// TIA Portal V21 export
// export: Created 2026-10-09T20:27:00.7380612Z, ExportSetting WithDefaults, DisplayName Totally Integrated Automation Portal, DisplayVersion V21, DisplayName STEP 7 Professional, DisplayVersion V21, DisplayName STEP 7 Safety, DisplayVersion V21, DisplayName Tech WebApplication, DisplayVersion V21, DisplayName WinCC Basic/Comfort/Advanced, DisplayVersion V21, DisplayName WinCC Unified, DisplayVersion V21
FUNCTION_BLOCK "FB_2_Filling"   // FB3, FBD
TITLE = Filling process
{ S7_Optimized_Access := 'TRUE' }
VERSION : 0.1
// stored: AutoNumber true, IsIECCheckEnabled false, IsRetainMemResEnabled false, MemoryReserve 100, SetENOAutomatically false, UDAEnableTagReadback false
   VAR_INPUT
      externalSignals : "typeSignals";   // signals from external model
   END_VAR
   VAR_IN_OUT
      model : "typeModel";   // model parameter
      operate : "typeOperate";   // application operation
      signals : "typeSignals";   // current signals from tank
      process : "typeProcess";   // current process information
      appSignals : "typeApp";
      hmiSignals : "typeHmi";
      errors : "typeError";   // error information
   END_VAR
   VAR
      statShiftingBottle : Bool;
      statShiftingTrigger : Bool;
      statShiftingTimer : Int;
      statHmiBottleLevel : Real;   // parameter for HMI to show current bottle level
      statHmiDoShift : Bool;   // trigger for HMI to shift bottles
      statHmiFaultyBottle : Bool;   // trigger for HMI for faulty bottle
      statBatchIdOld { ExternalAccessible := 'False'; ExternalVisible := 'False'; ExternalWritable := 'False'} : UDInt := 0;   // helper when batchID changed
      statFillingTankTrigger : Bool;
      statStartCounter { ExternalAccessible := 'False'; ExternalVisible := 'False'; ExternalWritable := 'False'} : Bool;
      statProducedStart { ExternalAccessible := 'False'; ExternalVisible := 'False'; ExternalWritable := 'False'} : UDInt;
      statProducedEnd { ExternalAccessible := 'False'; ExternalVisible := 'False'; ExternalWritable := 'False'} : UDInt;
      statSizeBatchID : USInt;
      statSizeNumberProduced : USInt;
      statStringBatchID : String;
      statStringProductID : String;
   END_VAR
   VAR_TEMP
      tempBottleMaxLevel : Real;
      tempTimerFinished : Bool;
      tempTimeOutput : Time;
      tempCurrentTime : DTL;
      tempTimeRet : Int;
   END_VAR
   VAR_TEMP   // added for the SCL form of the ladder/FBD networks
      _w1 : Bool;
      _w2 : Bool;
   END_VAR
BEGIN

REGION Network 1: Calculation of params
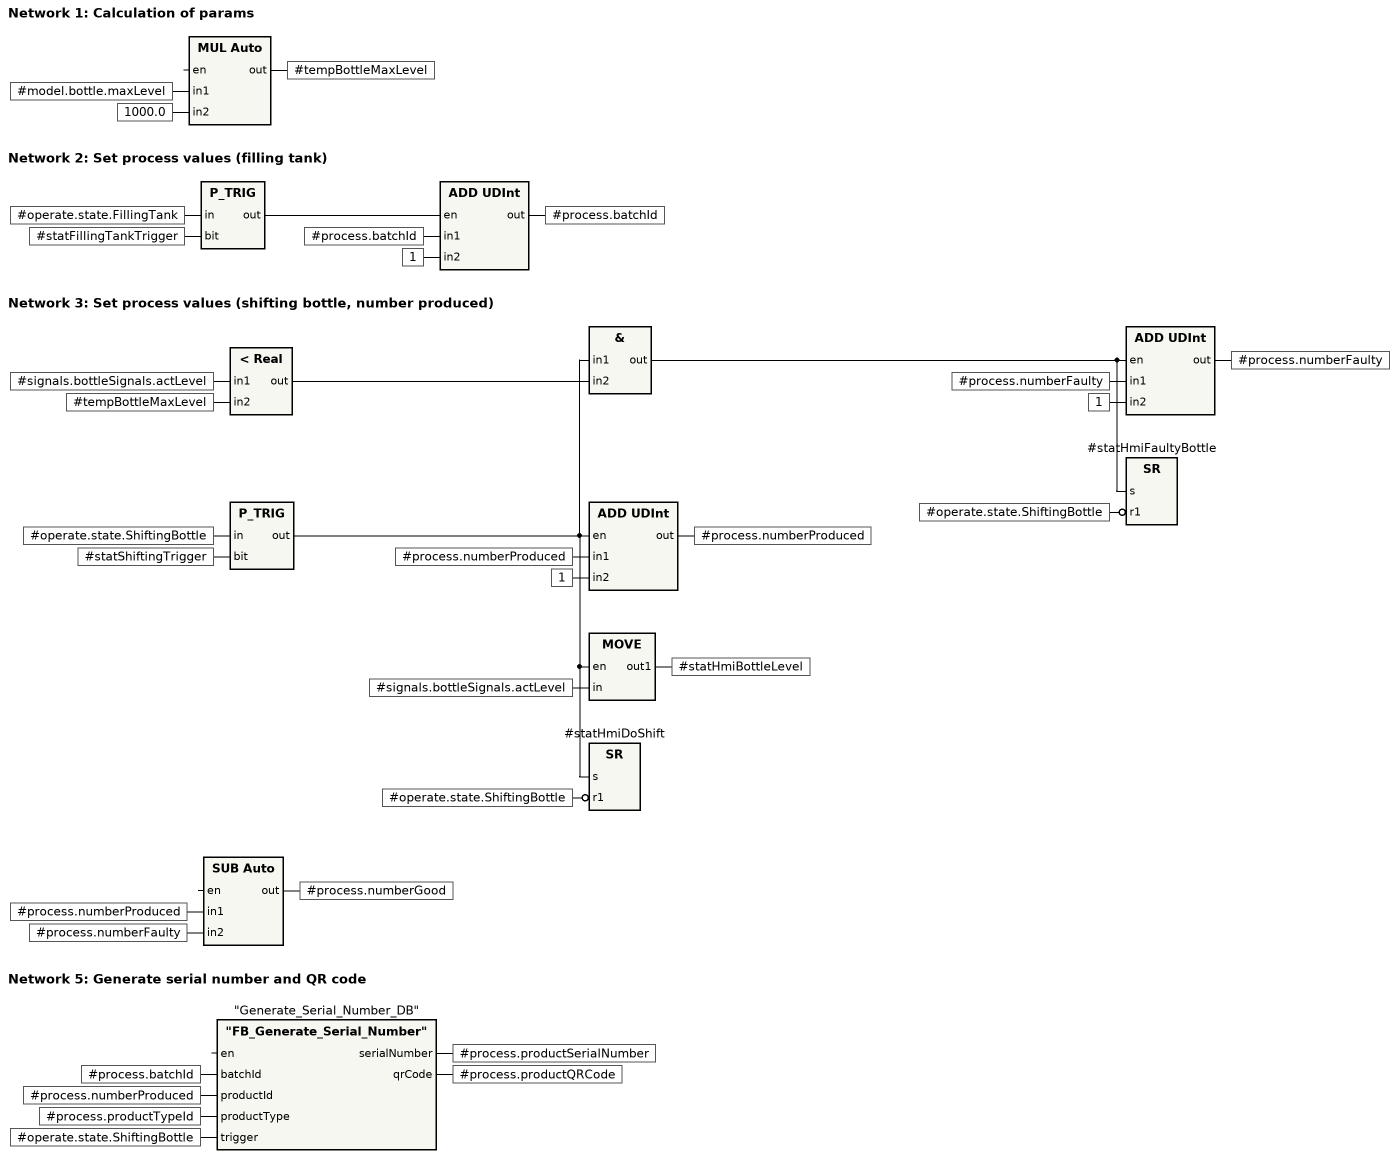
   #tempBottleMaxLevel := #model.bottle.maxLevel * 1000.0;
END_REGION

REGION Network 2: Set process values (filling tank)
   #_w1 := #operate.state.FillingTank AND NOT #statFillingTankTrigger;   // rising edge
   #statFillingTankTrigger := #operate.state.FillingTank;
   IF #_w1 THEN #process.batchId := #process.batchId + 1; END_IF;
END_REGION

REGION Network 3: Set process values (shifting bottle, number produced)
   #_w1 := #operate.state.ShiftingBottle AND NOT #statShiftingTrigger;   // rising edge
   #statShiftingTrigger := #operate.state.ShiftingBottle;
   IF #_w1 THEN #process.numberProduced := #process.numberProduced + 1; END_IF;
   #_w2 := #_w1 AND (#signals.bottleSignals.actLevel < #tempBottleMaxLevel);
   IF #_w2 THEN
       #process.numberFaulty := #process.numberFaulty + 1;
       #statHmiFaultyBottle := TRUE;   // SR flip-flop
   END_IF;
   IF NOT #operate.state.ShiftingBottle THEN #statHmiFaultyBottle := FALSE; END_IF;
   IF #_w1 THEN
       #statHmiBottleLevel := #signals.bottleSignals.actLevel;
       #statHmiDoShift := TRUE;   // SR flip-flop
   END_IF;
   IF NOT #operate.state.ShiftingBottle THEN #statHmiDoShift := FALSE; END_IF;
   #process.numberGood := #process.numberProduced - #process.numberFaulty;
END_REGION

REGION Network 4 (SCL): Set process values (product type ID, name)
   // 1 'Sparkling water'
   // 2 'Medium water'
   // 3 'Still water'
   IF #process.batchId <> #statBatchIdOld THEN

       IF #process.batchId = 1 THEN
           #process.productTypeId := 1;
       ELSE
           IF #process.productTypeId = 3 THEN
               #process.productTypeId := 1;
           ELSE
               #process.productTypeId := #process.productTypeId + 1;
           END_IF;
       END_IF;

       CASE #process.productTypeId OF
           1:  
               #process.productTypeName := 'Sparkling water';
           2:
               #process.productTypeName := 'Medium water';
           3:
               #process.productTypeName := 'Still water';
           ELSE
               #process.productTypeName := 'Undefined';
       END_CASE;

       #statBatchIdOld := #process.batchId;

   END_IF;
END_REGION

REGION Network 5: Generate serial number and QR code
   "Generate_Serial_Number_DB"(batchId := #process.batchId,   // "FB_Generate_Serial_Number"
                           productId := #process.numberProduced,
                           productType := #process.productTypeId,
                           trigger := #operate.state.ShiftingBottle,
                           serialNumber => #process.productSerialNumber,
                           qrCode => #process.productQRCode);
END_REGION

REGION Network 6 (SCL): Calculate production speed (pcs/h)
   // NOT WORKING currently
   // --> fix values as defined in GDB.process.speedActual


   (*

   // get current date
   #tempTimeRet := RD_LOC_T(#tempCurrentTime);  // get local time (DTL)

   // start counting every hour
   IF (#tempCurrentTime.MINUTE = 0 AND #tempCurrentTime.SECOND = 0) THEN
       #statStartCounter := true;
       #statProducedStart := #process.numberProduced;
   END_IF;

   "IEC_Timer_0_DB".TON(IN := #statStartCounter,
                        PT := T#59m_30s,
                        Q => #tempTimerFinished,
                        ET => #tempTimeOutput);

   IF #tempTimerFinished THEN
       #statStartCounter := false;
       #statProducedEnd := #process.numberProduced;
       IF #statProducedEnd > #statProducedStart THEN
           #process.speedActual := #statProducedEnd - #statProducedStart;
       ELSE
           #process.speedActual := 4294967295 - #statProducedStart + #statProducedEnd;
       END_IF;
   END_IF;

   *)
END_REGION

REGION Network 7 (SCL): Generate produt ID (batchID.numberProduced)
   IF #operate.state.ShiftingBottle THEN

       "FC_2_GetStringSizeOfNumber"(number := #process.batchId,
                                    stringSize => #statSizeBatchID);

       "FC_2_GetStringSizeOfNumber"(number := #process.numberProduced,
                                    stringSize => #statSizeNumberProduced);

       VAL_STRG(IN := #process.batchId,
                SIZE := #statSizeBatchID,
                PREC := 0,
                FORMAT := 0,
                P := 1,
                OUT => #statStringBatchID);

       VAL_STRG(IN := #process.numberProduced,
                SIZE := #statSizeNumberProduced,
                PREC := 0,
                FORMAT := 0,
                P := 1,
                OUT => #statStringProductID);

       #process.productId := CONCAT(
                                    IN1 := #statStringBatchID,
                                    IN2 := '.',
                                    IN3 := #statStringProductID
       );
   END_IF;
END_REGION

REGION Network 8 (SCL): Set cycle time
   CASE #operate.machineState OF
       "STATE_FILL_TANK":
           #model.cycleTime := 0.001;
       "STATE_HEAT_TANK":
           #model.cycleTime := 0.001;
       ELSE
           #model.cycleTime := 0.005;
   END_CASE;
END_REGION

REGION Network 9: Simulation (fill tank / heat tank / fill bottle)
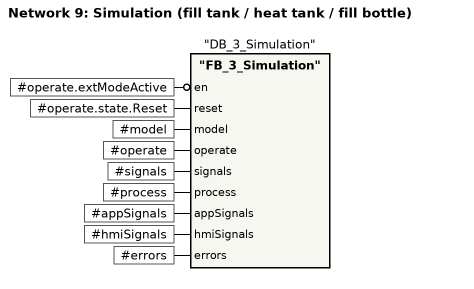
   IF NOT #operate.extModeActive THEN
       "DB_3_Simulation"(reset := #operate.state.Reset,   // "FB_3_Simulation"
                         model := #model,
                         operate := #operate,
                         signals := #signals,
                         process := #process,
                         appSignals := #appSignals,
                         hmiSignals := #hmiSignals,
                         errors := #errors);
   END_IF;
END_REGION

REGION Network 10 (SCL): Reset process parameter
   IF #operate.state.Reset THEN
       #process.batchId := 0;
       #process.numberFaulty := 0;
       #process.numberGood := 0;
       #process.numberProduced := 0;

       #process.productId := '';
       #process.productSerialNumber := '';
       #process.productTypeName := '';
       #process.productQRCode := 0;
       #process.productTypeId := 0;

       #process.speedActual := 0;
       #process.speedTarget := 0;

       #statHmiBottleLevel := 0.0;
       #signals.energySignals.energyConsumptionFillingBottles := 0.0;
       #signals.energySignals.energyConsumptionFillingTank := 0.0;
       #signals.energySignals.energyConsumptionHeatingTank := 0.0;
       #signals.energySignals.waterConsumptionFillingTank := 0.0;
       #signals.energySignals.gasConsumptionHeatingTank := 0.0;

   END_IF;
END_REGION
END_FUNCTION_BLOCK
